(* CODESYS project P_State.xml

Project tree, tasks and I/O mapping:
*)

// P_State
PROPERTY PRIVATE P_State : E_AlarmState
END_PROPERTY
